(* IEC 61131-3 sources: traffic-lights/PLC_TrafficLights/Class/_OpenSSL (part 2) *)

	FUNCTION __CDECL VIRTUAL GLOBAL CRYPTO_add_lock
		VAR_INPUT
			pointer 	: ^DINT;
			amount 	: DINT;
			t 	: DINT;
			file 	: ^void;
			line 	: DINT;
		END_VAR
		VAR_OUTPUT
			RetVal (EAX) 	: DINT;
		END_VAR;

	FUNCTION GLOBAL TAB RetVal;
				//! <Function Comment="X509_LOOKUP_file is a certificate lookup method to use with X509_STORE, provided by OpenSSL library.&#13;&#10;&#13;&#10;The X509_LOOKUP_file method loads all the certificates or CRLs present in a file into memory at the time the file is added as a lookup source.&#13;&#10;&#13;&#10;File format is ASCII text which contains concatenated PEM certificates and CRLs.&#13;&#10;&#13;&#10;This method should be used by applications which work with a small set of CAs.&#13;&#10;&#13;&#10;See also www.openssl.org/docs/man1.1.0/crypto/X509_LOOKUP_file.html&#13;&#10;and       www.umich.edu/~x509/ssleay/x509_lookup.html&#13;&#10;and       www.umich.edu/~x509/ssleay/x509_store.html" Name="X509_LOOKUP_file"/>
	FUNCTION __CDECL VIRTUAL GLOBAL X509_LOOKUP_file
		VAR_OUTPUT
			RetAddr (EAX) 	: ^void;			//! <Variable Comment="X509_LOOKUP_file() returns a X509_LOOKUP_METHOD pointer to the static method x509_file_lookup(). &#13;&#10;This function is useful to call when you want to add a method to a stack of methods you are using. &#13;&#10;See X509_STORE documentation for more on this." Name="X509_LOOKUP_file.RetAddr"/>
		END_VAR;
				//! <Function Comment="Issues arbitrary control commands.&#13;&#10;&#13;&#10;See also www.openssl.org/docs/manmaster/man3/X509_LOOKUP_meth_set_get_by_fingerprint.html" Name="X509_LOOKUP_ctrl"/>
	FUNCTION __CDECL VIRTUAL GLOBAL X509_LOOKUP_ctrl
		VAR_INPUT
			ctx 	: ^void;			//! <Variable Comment="Pointer to X509_LOOKUP structure." Name="X509_LOOKUP_ctrl.ctx"/>
			cmd 	: DINT;			//! <Variable Comment="An arbitrary integer that defines some operation." Name="X509_LOOKUP_ctrl.cmd"/>
			argc 	: ^void;			//! <Variable Comment="Pointer to an array of characters.&#13;&#10;How argc and argl are used depends entirely on the control function." Name="X509_LOOKUP_ctrl.argc"/>
			argl 	: DINT;			//! <Variable Comment="Arbitrary integer.&#13;&#10;How argc and argl are used depends entirely on the control function." Name="X509_LOOKUP_ctrl.argl"/>
			retv 	: ^pVoid;			//! <Variable Comment="NULL or pointer to pointer to a location where any return data should be written to." Name="X509_LOOKUP_ctrl.retv"/>
		END_VAR
		VAR_OUTPUT
			RetVal (EAX) 	: DINT;			//! <Variable Comment="Returns -1 if no method table was found.&#13;&#10;              1 if no lookup method was found.&#13;&#10;" Name="X509_LOOKUP_ctrl.RetVal"/>
		END_VAR;
				//! <Function Comment="The X509_verify_cert() function attempts to discover and validate a certificate chain based on parameters in &lt;ctx&gt;. &#13;&#10;A complete description of the process is contained in the verify manual page. &#13;&#10;&#13;&#10;See also www.openssl.org/docs/manmaster/man3/X509_verify_cert.html" Name="X509_verify_cert"/>
	FUNCTION __CDECL VIRTUAL GLOBAL X509_verify_cert
		VAR_INPUT
			ctx 	: ^void;			//! <Variable Comment="Pointer to a context (X509_STORE_CTX structure)." Name="X509_verify_cert.ctx"/>
		END_VAR
		VAR_OUTPUT
			RetVal (EAX) 	: DINT;			//! <Variable Comment="If a complete chain can be built and validated this function returns 1, otherwise it return zero, in exceptional circumstances it can also return a negative code." Name="X509_verify_cert.RetVal"/>
		END_VAR;
				//! <Function Comment="X509_NAME_oneline() prints an ASCII version of &lt;a&gt; to &lt;buf&gt;. If &lt;buf&gt; is NULL then a buffer is dynamically allocated and returned, and &lt;size&gt; is ignored. &#13;&#10;Otherwise, at most &lt;size&gt; bytes will be written, including the ending &apos;\0&apos;, and &lt;buf&gt; is returned.&#13;&#10;&#13;&#10;NOTES&#13;&#10;X509_NAME_oneline() is a legacy function which produces a nonstandard output form, it doesn&apos;t handle multi character fields and has various quirks and inconsistencies. &#13;&#10;Its use is strongly discouraged in new applications.&#13;&#10;&#13;&#10;See also www.openssl.org/docs/man1.0.2/crypto/X509_NAME_oneline.html" Name="X509_NAME_oneline"/>
	FUNCTION __CDECL VIRTUAL GLOBAL X509_NAME_oneline
		VAR_INPUT
			a 	: ^void;			//! <Variable Comment="Pointer to a X509_NAME structure." Name="X509_NAME_oneline.a"/>
			buf 	: ^void;			//! <Variable Comment="Pointer to an output buffer or NULL (*char)." Name="X509_NAME_oneline.buf"/>
			size 	: DINT;			//! <Variable Comment="Output buffer size." Name="X509_NAME_oneline.size"/>
		END_VAR
		VAR_OUTPUT
			RetAddr (EAX) 	: ^void;			//! <Variable Comment="Pointer to the output buffer (*char)." Name="X509_NAME_oneline.RetAddr"/>
		END_VAR;
				//! <Function Comment="Internally loading of CRLs is implemented via function X509_load_crl_file. &#13;&#10;The function supports parameter &lt;typ&gt;, which can be one of constants FILETYPE_PEM, FILETYPE_ASN1 and FILETYPE_DEFAULT. &#13;&#10;It loads CRLs from specified &lt;file&gt; into memory cache of X509_STORE objects which given &lt;ctx&gt; parameter is associated with.&#13;&#10;&#13;&#10;See also www.openssl.org/docs/man1.1.0/crypto/X509_load_crl_file.html" Name="X509_load_crl_file"/>
	FUNCTION __CDECL VIRTUAL GLOBAL X509_load_crl_file
		VAR_INPUT
			ctx 	: ^void;			//! <Variable Comment="Pointer to X509_LOOKUP structure." Name="X509_load_crl_file.ctx"/>
			file 	: ^void;			//! <Variable Comment="Specifies the file to read from." Name="X509_load_crl_file.file"/>
			typ 	: DINT;			//! <Variable Comment="Can be one of constants FILETYPE_PEM, FILETYPE_ASN1 and FILETYPE_DEFAULT." Name="X509_load_crl_file.typ"/>
		END_VAR
		VAR_OUTPUT
			RetVal (EAX) 	: DINT;			//! <Variable Comment="Returns number of objects loaded from &lt;file&gt; or 0 in case of error." Name="X509_load_crl_file.RetVal"/>
		END_VAR;
				//! <Function Comment="X509_STORE_CTX_new() returns a newly initialised X509_STORE_CTX structure.&#13;&#10;&#13;&#10;NOTES&#13;&#10;The certificates and CRLs in a store are used internally and should not be freed up until after the associated X509_STORE_CTX is freed.&#13;&#10;&#13;&#10;BUGS&#13;&#10;The certificates and CRLs in a context are used internally and should not be freed up until after the associated X509_STORE_CTX is freed. &#13;&#10;Copies should be made, or reference counts increased instead.&#13;&#10;&#13;&#10;See also www.openssl.org/docs/man1.1.0/crypto/X509_STORE_CTX_new.html" Name="X509_STORE_CTX_new"/>
	FUNCTION __CDECL VIRTUAL GLOBAL X509_STORE_CTX_new
		VAR_OUTPUT
			RetAddr (EAX) 	: ^void;			//! <Variable Comment="Returns an newly allocated context (Pointer to X509_STORE_CTX structure) or &#13;&#10;NULL if an error occurred." Name="X509_STORE_CTX_new.RetAddr"/>
		END_VAR;
				//! <Function Comment="X509_STORE_CTX_free() completely frees up &lt;ctx&gt;. After this call &lt;ctx&gt; is no longer valid. &#13;&#10;If &lt;ctx&gt; is NULL nothing is done.&#13;&#10;&#13;&#10;See also www.openssl.org/docs/man1.1.0/crypto/X509_STORE_CTX_new.html" Name="X509_STORE_CTX_free"/>
	FUNCTION __CDECL VIRTUAL GLOBAL X509_STORE_CTX_free
		VAR_INPUT
			ctx 	: ^void;			//! <Variable Comment="Pointer to X509_STORE_CTX structure holding a context." Name="X509_STORE_CTX_free.ctx"/>
		END_VAR;
				//! <Function Comment="X509_STORE_CTX_init() sets up &lt;ctx&gt; for a subsequent verification operation. &#13;&#10;It must be called before each call to X509_verify_cert(), i.e. a &lt;ctx&gt; is only good for one call to X509_verify_cert(). &#13;&#10;If you want to verify a second certificate with the same &lt;ctx&gt; then you must call X509_STORE_CTX_cleanup() and then X509_STORE_CTX_init() again before the second call to X509_verify_cert(). &#13;&#10;The trusted certificate store is set to &lt;store&gt;, the end entity certificate to be verified is set to &lt;x509&gt; and a set of additional certificates (which will be untrusted but may be used to build the chain) in &lt;chain&gt;. &#13;&#10;Any or all of the &lt;store&gt;, &lt;x509&gt; and &lt;chain&gt; parameters can be NULL.&#13;&#10;&#13;&#10;See also www.openssl.org/docs/man1.1.0/crypto/X509_STORE_CTX_new.html" Name="X509_STORE_CTX_init"/>
	FUNCTION __CDECL VIRTUAL GLOBAL X509_STORE_CTX_init
		VAR_INPUT
			ctx 	: ^void;			//! <Variable Comment="Pointer to X509_STORE_CTX structure." Name="X509_STORE_CTX_init.ctx"/>
			store 	: ^void;			//! <Variable Comment="Pointer to X509_STORE structure or NULL" Name="X509_STORE_CTX_init.store"/>
			x509 	: ^void;			//! <Variable Comment="Pointer to X509 structure or NULL." Name="X509_STORE_CTX_init.x509"/>
			chain 	: ^void;			//! <Variable Comment="Pointer to STACK_OF(X509) or NULL." Name="X509_STORE_CTX_init.chain"/>
		END_VAR
		VAR_OUTPUT
			RetVal (EAX) 	: DINT;			//! <Variable Comment="Returns 1 for success or 0 if an error occurred." Name="X509_STORE_CTX_init.RetVal"/>
		END_VAR;
				//! <Function Comment="Returns the issuer name of certificate &lt;a&gt;. The returned value is an internal pointer which MUST NOT be freed.&#13;&#10;&#13;&#10;See also www.openssl.org/docs/man1.1.0/crypto/X509_get_subject_name.html" Name="X509_get_issuer_name"/>
	FUNCTION __CDECL VIRTUAL GLOBAL X509_get_issuer_name
		VAR_INPUT
			a 	: ^void;			//! <Variable Comment="Pointer to X509 structure holding a certificate." Name="X509_get_issuer_name.a"/>
		END_VAR
		VAR_OUTPUT
			RetAddr (EAX) 	: ^void;			//! <Variable Comment="Returns an X509_NAME pointer." Name="X509_get_issuer_name.RetAddr"/>
		END_VAR;
				//! <Function Comment="X509_LOOKUP_hash_dir is a certificate lookup method to use with X509_STORE, provided by OpenSSL library. &#13;&#10;X509_LOOKUP_hash_dir is a more advanced method, which loads certificates and CRLs on demand, and caches them in memory once they are loaded.&#13;&#10;&#13;&#10;See also www.openssl.org/docs/man1.1.0/crypto/X509_LOOKUP_hash_dir.html&#13;&#10;and       http://www.umich.edu/~x509/ssleay/x509_store.html" Name="X509_LOOKUP_hash_dir"/>
	FUNCTION __CDECL VIRTUAL GLOBAL X509_LOOKUP_hash_dir
		VAR_OUTPUT
			RetVal (EAX) 	: ^void;			//! <Variable Comment="Returns 1 on success or 0 on error. " Name="X509_LOOKUP_hash_dir.RetVal"/>
		END_VAR;
				//! <Function Comment="Sets the default values for the corresponding values used in certificate chain validation. &#13;&#10;Their behavior is documented in the corresponding X509_VERIFY_PARAM manual pages, e.g., X509_VERIFY_PARAM_set_depth(3).&#13;&#10;&#13;&#10;See also www.openssl.org/docs/manmaster/man3/X509_STORE_set_flags.html" Name="X509_STORE_set_flags"/>
	FUNCTION __CDECL VIRTUAL GLOBAL X509_STORE_set_flags
		VAR_INPUT
			ctx 	: ^void;			//! <Variable Comment="Pointer to X509_STORE structure.&#13;&#10;&#13;&#10;The X509_STORE structure is intended to be a consolidated mechanism for holding information about X.509 certificates and CRLs, and constructing and validating chains of certificates terminating in trusted roots. &#13;&#10;It admits multiple lookup mechanisms and efficient scaling performance with large numbers of certificates, and a great deal of flexibility in how validation and policy checks are performed." Name="X509_STORE_set_flags.ctx"/>
			flags 	: UDINT;			//! <Variable Comment="Flag values to set." Name="X509_STORE_set_flags.flags"/>
		END_VAR
		VAR_OUTPUT
			RetVal (EAX) 	: DINT;			//! <Variable Comment="Always returns 1, indicating success." Name="X509_STORE_set_flags.RetVal"/>
		END_VAR;
				//! <Function Comment="Adds the X509_LOOKUP_METHOD &lt;a&gt; to the stack &lt;v&gt;-&gt;get_cert_methods after creating an X509_LOOKUP that contains it as a subfield. &#13;&#10;It returns a pointer to the new X509_LOOKUP structure or NULL on error.&#13;&#10;&#13;&#10;X509_STORE_new() creates an empty X509_STORE structure, which contains no information about trusted certificates or where such certificates are located on disk, and is generally not usable. &#13;&#10;Normally, trusted certificates will be added to the X509_STORE to prepare it for use, via mechanisms such as X509_STORE_add_lookup() and X509_LOOKUP_file(), or PEM_read_bio_X509_AUX() &#13;&#10;and X509_STORE_add_cert(). &#13;&#10;CRLs can also be added, and many behaviors configured as desired.&#13;&#10;&#13;&#10;See also http://www.umich.edu/~x509/ssleay/x509_store.html&#13;&#10;" Name="X509_STORE_add_lookup"/>
	FUNCTION __CDECL VIRTUAL GLOBAL X509_STORE_add_lookup
		VAR_INPUT
			v 	: ^void;			//! <Variable Comment="Pointer to X509_STORE structure." Name="X509_STORE_add_lookup.v"/>
			a 	: ^void;			//! <Variable Comment="Pointer to X509_LOOKUP_METHOD structure holding a lookup method." Name="X509_STORE_add_lookup.a"/>
		END_VAR
		VAR_OUTPUT
			RetAddr (EAX) 	: ^void;			//! <Variable Comment="Returns a pointer to the new X509_LOOKUP structure or NULL on error." Name="X509_STORE_add_lookup.RetAddr"/>
		END_VAR;
				//! <Function Comment="X509_STORE_set_default_paths() is somewhat misnamed, in that it does not set what default paths should be used for loading certificates. &#13;&#10;Instead, it loads certificates into the X509_STORE from the hardcoded default paths.&#13;&#10;&#13;&#10;See also www.openssl.org/docs/man1.1.1/man3/X509_STORE_set_default_paths.html&#13;&#10;and       http://www.umich.edu/~x509/ssleay/x509_store.html" Name="X509_STORE_set_default_paths"/>
	FUNCTION __CDECL VIRTUAL GLOBAL X509_STORE_set_default_paths
		VAR_INPUT
			ctx 	: ^void;			//! <Variable Comment="Pointer to X509_STORE structure." Name="X509_STORE_set_default_paths.ctx"/>
		END_VAR
		VAR_OUTPUT
			RetVal (EAX) 	: DINT;			//! <Variable Comment="Returns 1 on success or 0 on failure." Name="X509_STORE_set_default_paths.RetVal"/>
		END_VAR;
				//! <Function Comment="Is used to retrieve application specific data. Returns the application data or 0 on failure. &#13;&#10;0 may also be valid application data but currently it can only fail if given an invalid &lt;idx&gt; parameter.&#13;&#10;&#13;&#10;See also www.openssl.org/docs/man1.0.2/crypto/X509_STORE_CTX_get_ex_data.html&#13;&#10;and       www.openssl.org/docs/man1.0.2/crypto/RSA_get_ex_new_index.html" Name="X509_STORE_CTX_get_ex_data"/>
	FUNCTION __CDECL VIRTUAL GLOBAL X509_STORE_CTX_get_ex_data
		VAR_INPUT
			ctx 	: ^void;			//! <Variable Comment="Pointer to X509_STORE_CTX structure." Name="X509_STORE_CTX_get_ex_data.ctx"/>
			idx 	: DINT;			//! <Variable Comment="Index retrieved by RSA_get_ex_new_index()." Name="X509_STORE_CTX_get_ex_data.idx"/>
		END_VAR
		VAR_OUTPUT
			RetAddr (EAX) 	: ^void;			//! <Variable Comment="Pointer to the retrieved application data or NULL on failure.&#13;&#10;Since the application data can be anything at all it is passed and retrieved as a void * type." Name="X509_STORE_CTX_get_ex_data.RetAddr"/>
		END_VAR;
				//! <Function Comment="Is used to set application specific data, the data is supplied in the &lt;data&gt; parameter and its precise meaning is up to the application.&#13;&#10;&#13;&#10;See also www.openssl.org/docs/man1.0.2/crypto/X509_STORE_CTX_get_ex_data.html&#13;&#10;and       www.openssl.org/docs/man1.0.2/crypto/RSA_get_ex_new_index.html" Name="X509_STORE_CTX_set_ex_data"/>
	FUNCTION __CDECL VIRTUAL GLOBAL X509_STORE_CTX_set_ex_data
		VAR_INPUT
			ctx 	: ^void;			//! <Variable Comment="Pointer to X509_STORE_CTX structure." Name="X509_STORE_CTX_set_ex_data.ctx"/>
			idx 	: DINT;			//! <Variable Comment="Index retrieved by RSA_get_ex_new_index()." Name="X509_STORE_CTX_set_ex_data.idx"/>
			data 	: ^void;			//! <Variable Comment="Pointer to the application data.&#13;&#10;Since the application data can be anything at all it is passed as a void * type." Name="X509_STORE_CTX_set_ex_data.data"/>
		END_VAR
		VAR_OUTPUT
			RetVal (EAX) 	: DINT;			//! <Variable Comment="Returns 1 on success or 0 on failure." Name="X509_STORE_CTX_set_ex_data.RetVal"/>
		END_VAR;
				//! <Function Comment="X509_STORE_CTX_get_error() returns the error code of &lt;ctx&gt;, see the ERROR CODES section for a full description of all error codes. &#13;&#10;&#13;&#10;This function is typically called after X509_verify_cert() has indicated an error or in a verification callback to determine the nature of an error.&#13;&#10;&#13;&#10;See also www.openssl.org/docs/man1.0.2/crypto/X509_STORE_CTX_get_error.html" Name="X509_STORE_CTX_get_error"/>
	FUNCTION __CDECL VIRTUAL GLOBAL X509_STORE_CTX_get_error
		VAR_INPUT
			ctx 	: ^void;			//! <Variable Comment="Pointer to X509_STORE_CTX structure." Name="X509_STORE_CTX_get_error.ctx"/>
		END_VAR
		VAR_OUTPUT
			RetVal (EAX) 	: DINT;			//! <Variable Comment="Returns X509_V_OK or an error code.&#13;&#10;&#13;&#10;See the class documentation for a list of error codes and messages." Name="X509_STORE_CTX_get_error.RetVal"/>
		END_VAR;
				//! <Function Comment="X509_STORE_CTX_get_current_cert() returns the certificate in &lt;ctx&gt; which caused the error or NULL if no certificate is relevant.&#13;&#10;&#13;&#10;This function is typically called after X509_verify_cert() has indicated an error or in a verification callback to determine the nature of an error.&#13;&#10;&#13;&#10;See also www.openssl.org/docs/man1.0.2/crypto/X509_STORE_CTX_get_error.html" Name="X509_STORE_CTX_get_current_cert"/>
	FUNCTION __CDECL VIRTUAL GLOBAL X509_STORE_CTX_get_current_cert
		VAR_INPUT
			ctx 	: ^void;			//! <Variable Comment="Pointer to X509_STORE_CTX structure." Name="X509_STORE_CTX_get_current_cert.ctx"/>
		END_VAR
		VAR_OUTPUT
			RetAddr (EAX) 	: ^void;			//! <Variable Comment="Returns a X509 pointer to the certificate which caused the error or NULL if no certificate is relevant to the error." Name="X509_STORE_CTX_get_current_cert.RetAddr"/>
		END_VAR;
				//! <Function Comment="X509_STORE_CTX_get_error_depth() returns the depth of the error. This is a non-negative integer representing where in the certificate chain the error occurred. &#13;&#10;If it is zero it occurred in the end entity certificate, one if it is the certificate which signed the end entity certificate and so on.&#13;&#10;&#13;&#10;This function is typically called after X509_verify_cert() has indicated an error or in a verification callback to determine the nature of an error.&#13;&#10;&#13;&#10;See also www.openssl.org/docs/man1.0.2/crypto/X509_STORE_CTX_get_error.html" Name="X509_STORE_CTX_get_error_depth"/>
	FUNCTION __CDECL VIRTUAL GLOBAL X509_STORE_CTX_get_error_depth
		VAR_INPUT
			ctx 	: ^void;			//! <Variable Comment="Pointer to X509_STORE_CTX structure." Name="X509_STORE_CTX_get_error_depth.ctx"/>
		END_VAR
		VAR_OUTPUT
			RetVal (EAX) 	: DINT;			//! <Variable Comment="Returns a non-negative error depth." Name="X509_STORE_CTX_get_error_depth.RetVal"/>
		END_VAR;
				//! <Function Comment="X509_verify_cert_error_string() returns a human readable error string for verification of error &lt;a&gt;." Name="X509_verify_cert_error_string"/>
	FUNCTION __CDECL VIRTUAL GLOBAL X509_verify_cert_error_string
		VAR_INPUT
			a 	: DINT;			//! <Variable Comment="Error number." Name="X509_verify_cert_error_string.a"/>
		END_VAR
		VAR_OUTPUT
			RetAddr (EAX) 	: ^void;			//! <Variable Comment="Returns a human readable error string for verification of error &lt;a&gt;." Name="X509_verify_cert_error_string.RetAddr"/>
		END_VAR;
				//! <Function Comment="i2d_PublicKey() encodes key &lt;a&gt; into DER format. It uses a key specific format or, if none is defined for that key type, PKCS#8 unencrypted PublicKeyInfo format.&#13;&#10;&#13;&#10;NOTES&#13;&#10;The EVP_PKEY structure passed to the function should have all the public key components present.&#13;&#10;&#13;&#10;The encoded data is in binary form and may contain embedded zeroes. Functions such as strlen() will not return the correct length of the encoded structure.&#13;&#10;&#13;&#10;See also www.openssl.org/docs/man1.1.0/crypto/i2d_PublicKey.html&#13;&#10;and       www.openssl.org/docs/man1.0.2/crypto/i2d_RSAPublicKey.html&#13;&#10;and       www.openssl.org/docs/manmaster/man3/i2d_RSA_PUBKEY.html" Name="i2d_PublicKey"/>
	FUNCTION __CDECL VIRTUAL GLOBAL i2d_PublicKey
		VAR_INPUT
			a 	: ^void;			//! <Variable Comment="Pointer to a EVP_PKEY structure holding the public key." Name="i2d_PublicKey.a"/>
			pp 	: ^pVoid;			//! <Variable Comment="Pointer to pointer to output buffer (i.e. **char).&#13;&#10;If &lt;pp&gt; is not NULL, the DER encoded data is written to the buffer at *&lt;pp&gt;, and *&lt;pp&gt; is incremented to point after the data just written.&#13;&#10;If *&lt;pp&gt; is NULL memory will be allocated for a buffer and the encoded data written to it. In this case *&lt;pp&gt; is not incremented and it points to the start of the data just written." Name="i2d_PublicKey.pp"/>
		END_VAR
		VAR_OUTPUT
			RetVal (EAX) 	: DINT;			//! <Variable Comment="Returns the number of bytes successfully encoded or a negative value if an error occurs. &#13;&#10;The error code can be obtained by calling ERR_get_error()." Name="i2d_PublicKey.RetVal"/>
		END_VAR;
				//! <Function Comment="EVP_PKEY_type() returns the type of key corresponding to the value &lt;typ&gt;. &#13;&#10;The type of a key can be obtained with EVP_PKEY_type(pkey-&gt;type). &#13;&#10;&#13;&#10;See also www.openssl.org/docs/man1.0.2/crypto/EVP_PKEY_type.html" Name="EVP_PKEY_type"/>
	FUNCTION __CDECL VIRTUAL GLOBAL EVP_PKEY_type
		VAR_INPUT
			typ 	: DINT;			//! <Variable Comment="Value retrieved with pkey-&gt;type." Name="EVP_PKEY_type.typ"/>
		END_VAR
		VAR_OUTPUT
			RetVal (EAX) 	: DINT;			//! <Variable Comment="The return value will be EVP_PKEY_RSA, EVP_PKEY_DSA, EVP_PKEY_DH or EVP_PKEY_EC for the corresponding key types or NID_undef if the key type is unassigned." Name="EVP_PKEY_type.RetVal"/>
		END_VAR;
				//! <Function Comment="Do not use this function in new code. It is provided purely for compatibility with legacy application code.&#13;&#10;This function is a wrapper around the corresponding standard realloc() function.&#13;&#10;&#13;&#10;See also www.openssl.org/docs/man1.1.0/crypto/CRYPTO_realloc.html&#13;&#10;and       http://man.openbsd.org/OpenBSD-6.1/OPENSSL_realloc.3" Name="CRYPTO_realloc"/>
	FUNCTION __CDECL VIRTUAL GLOBAL CRYPTO_realloc
		VAR_INPUT
			addr 	: ^void;			//! <Variable Comment="Pointer to a memory block previously allocated." Name="CRYPTO_realloc.addr"/>
			num 	: DINT;			//! <Variable Comment="New size for the memory block, in bytes." Name="CRYPTO_realloc.num"/>
			file 	: ^void;			//! <Variable Comment="The Structured Text __FILE__ parameter." Name="CRYPTO_realloc.file"/>
			line 	: DINT;			//! <Variable Comment="The Structured Text __LINE__ parameter." Name="CRYPTO_realloc.line"/>
		END_VAR
		VAR_OUTPUT
			RetAddr (EAX) 	: ^void;			//! <Variable Comment="Returns a void pointer to allocated memory or NULL on error." Name="CRYPTO_realloc.RetAddr"/>
		END_VAR;
				//! <Function Comment="BIO_ctrl() is a BIO &quot;control&quot; operation taking arguments of various types. &#13;&#10;This function is not normally called directly, various macros are used instead. &#13;&#10;The standard macros are described below, macros specific to a particular type of BIO are described in the specific BIOs manual page as well as any special features of the standard calls.&#13;&#10;&#13;&#10;A BIO is an I/O abstraction, it hides many of the underlying I/O details from an application. &#13;&#10;If an application uses a BIO for its I/O it can transparently handle SSL connections, unencrypted network connections and file I/O.&#13;&#10;&#13;&#10;See also www.openssl.org/docs/man1.0.2/crypto/BIO_ctrl.html&#13;&#10;and       www.openssl.org/docs/man1.0.2/crypto/BIO_get_read_request.html&#13;&#10;and       www.openssl.org/docs/man1.0.2/crypto/BIO_new_buffer_ssl_connect.html&#13;&#10;and       www.openssl.org/docs/man1.0.2/crypto/BIO_ctrl_reset_read_request.html&#13;&#10;and       www.openssl.org/docs/man1.0.2/crypto/BIO_f_buffer.html&#13;&#10;and       www.openssl.org/docs/man1.0.2/crypto/BIO_set_fd.html&#13;&#10;and       www.openssl.org/docs/man1.1.1/man7/bio.html" Name="BIO_ctrl"/>
	FUNCTION __CDECL VIRTUAL GLOBAL BIO_ctrl
		VAR_INPUT
			b 	: ^void;			//! <Variable Comment="Pointer to BIO structure." Name="BIO_ctrl.b"/>
			cmd 	: DINT;			//! <Variable Comment="Command code.&#13;&#10;E.g. BIO_C_MAKE_BIO_PAIR, BIO_C_DESTROY_BIO_PAIR, &#13;&#10;BIO_C_SHUTDOWN_WR, BIO_C_SET_WRITE_BUF_SIZE, BIO_C_GET_WRITE_BUF_SIZE, &#13;&#10;BIO_C_GET_WRITE_GUARANTEE, BIO_C_GET_READ_REQUEST,&#13;&#10;BIO_C_SET_SSL, BIO_C_GET_SSL,&#13;&#10;BIO_C_SSL_MODE,&#13;&#10;BIO_C_SET_SSL_RENEGOTIATE_BYTES,&#13;&#10;BIO_C_SET_SSL_RENEGOTIATE_TIMEOUT,&#13;&#10;BIO_C_SET_SSL_NUM_RENEGOTIATES,&#13;&#10;BIO_C_DO_STATE_MACHINE ........" Name="BIO_ctrl.cmd"/>
			larg 	: DINT;			//! <Variable Comment="The meaning of &lt;larg&gt; depends on parameter &lt;cmd&gt;." Name="BIO_ctrl.larg"/>
			parg 	: ^void;			//! <Variable Comment="The meaning of &lt;parg&gt; depends on parameter &lt;cmd&gt;." Name="BIO_ctrl.parg"/>
		END_VAR
		VAR_OUTPUT
			RetVal (EAX) 	: DINT;			//! <Variable Comment="The meaning of &lt;RetVal&gt; depends on parameter &lt;cmd&gt;." Name="BIO_ctrl.RetVal"/>
		END_VAR;
				//! <Function Comment="BIO_s_mem() returns the memory BIO method function.&#13;&#10;A memory BIO is a source/sink BIO which uses memory for its I/O." Name="BIO_s_mem"/>
	FUNCTION __CDECL VIRTUAL GLOBAL BIO_s_mem
		VAR_OUTPUT
			RetAddr (EAX) 	: ^void;			//! <Variable Comment="Returns a BIO_METHOD pointer to the memory BIO method function." Name="BIO_s_mem.RetAddr"/>
		END_VAR;
				//! <Function Comment="BIO_s_file() returns the BIO file method. As its name implies it is a wrapper round the stdio FILE structure and it is a source/sink BIO.&#13;&#10;&#13;&#10;See also www.openssl.org/docs/man1.0.2/crypto/BIO_s_file.html" Name="BIO_s_file"/>
	FUNCTION __CDECL VIRTUAL GLOBAL BIO_s_file
		VAR_OUTPUT
			RetAddr (EAX) 	: ^void;			//! <Variable Comment="Returns a BIO_METHOD pointer to the BIO file method." Name="BIO_s_file.RetAddr"/>
		END_VAR;
				//! <Function Comment="X509_get_ext() operates on the extensions of certificate &lt;x&gt;. It is otherwise identical to X509v3_get_ext().&#13;&#10;&#13;&#10;X509v3_get_ext() retrieves extension &lt;loc&gt; from &lt;x&gt;. The index &lt;loc&gt; can take any value from 0 to X509_get_ext_count(&lt;x&gt;) - 1. &#13;&#10;The returned extension is an internal pointer which must not be freed up by the application.&#13;&#10;&#13;&#10;See also www.openssl.org/docs/man1.1.0/crypto/X509_get_ext.html" Name="X509_get_ext"/>
	FUNCTION __CDECL VIRTUAL GLOBAL X509_get_ext
		VAR_INPUT
			x 	: ^void;			//! <Variable Comment="Pointer to X509 structure holding a certificate." Name="X509_get_ext.x"/>
			loc 	: DINT;			//! <Variable Comment="Any value from 0 to X509_get_ext_count(&lt;x&gt;) - 1. " Name="X509_get_ext.loc"/>
		END_VAR
		VAR_OUTPUT
			RetAddr (EAX) 	: ^void;			//! <Variable Comment="Returns an X509_EXTENSION pointer or NULL if an error occurs." Name="X509_get_ext.RetAddr"/>
		END_VAR;
				//! <Function Comment="The function EVP_PKEY_cmp() compares the public key components and parameters (if present) of keys &lt;a&gt; and &lt;b&gt;.&#13;&#10;&#13;&#10;See also www.openssl.org/docs/man1.0.2/crypto/EVP_PKEY_cmp.html" Name="EVP_PKEY_cmp"/>
	FUNCTION __CDECL VIRTUAL GLOBAL EVP_PKEY_cmp
		VAR_INPUT
			a 	: ^void;			//! <Variable Comment="EVP_PKEY pointer to first key." Name="EVP_PKEY_cmp.a"/>
			b 	: ^void;			//! <Variable Comment="EVP_PKEY pointer to second key." Name="EVP_PKEY_cmp.b"/>
		END_VAR
		VAR_OUTPUT
			RetVal (EAX) 	: DINT;			//! <Variable Comment="Returns &#13;&#10;1 if the keys match, &#13;&#10;0 if they don&apos;t match, &#13;&#10;-1 if the key types are different and &#13;&#10;-2 if the operation is not supported." Name="EVP_PKEY_cmp.RetVal"/>
		END_VAR;
				//! <Function Comment="The EVP_PKEY_new() function allocates an empty EVP_PKEY structure which is used by OpenSSL to store private keys.&#13;&#10;EVP_PKEY_free() frees up the private key key.&#13;&#10;&#13;&#10;NOTES&#13;&#10;The EVP_PKEY structure is used by various OpenSSL functions which require a general private key without reference to any particular algorithm.&#13;&#10;&#13;&#10;The structure returned by EVP_PKEY_new() is empty. To add a private key to this empty structure the functions described in EVP_PKEY_set1_RSA should be used.&#13;&#10;&#13;&#10;See also www.openssl.org/docs/man1.0.2/crypto/EVP_PKEY_new.html" Name="EVP_PKEY_new"/>
	FUNCTION __CDECL VIRTUAL GLOBAL EVP_PKEY_new
		VAR_OUTPUT
			RetAddr (EAX) 	: ^void;			//! <Variable Comment="Returns either a pointer to the newly allocated EVP_PKEY structure of NULL if an error occurred." Name="EVP_PKEY_new.RetAddr"/>
		END_VAR;
				//! <Function Comment="The function ASN1_TIME_set() sets the ASN1_TIME structure &lt;sx&gt; to the time represented by the time_t value &lt;tx&gt;. &#13;&#10;If &lt;sx&gt; is NULL a new ASN1_TIME structure is allocated and returned.&#13;&#10;&#13;&#10;See also www.openssl.org/docs/man1.0.2/crypto/ASN1_TIME_set.html" Name="ASN1_TIME_set"/>
	FUNCTION __CDECL VIRTUAL GLOBAL ASN1_TIME_set
		VAR_INPUT
			sx 	: ^void;			//! <Variable Comment="Pointer to ASN1_TIME structure.&#13;&#10;&lt;sx&gt; must satisfy the ASN1_TIME format mandated by RFC 5280, i.e., its format must be either YYMMDDHHMMSSZ or YYYYMMDDHHMMSSZ (it&apos;s a literal Z at the end, meaning &quot;Zulu&quot;).&#13;&#10;" Name="ASN1_TIME_set.sx"/>
			tx 	: DINT;			//! <Variable Comment="Number of seconds since the start of the Unix epoch: midnight UTC of January 1, 1970 (not counting leap seconds)." Name="ASN1_TIME_set.tx"/>
		END_VAR
		VAR_OUTPUT
			RetAddr (EAX) 	: ^void;			//! <Variable Comment="Returns a pointer to an ASN1_TIME structure or NULL if an error occurred." Name="ASN1_TIME_set.RetAddr"/>
		END_VAR;
				//! <Function Comment="X509_CRL_sign() signs CRLs (Certificate Revocation Lists).&#13;&#10;&#13;&#10;See also www.openssl.org/docs/man1.1.0/crypto/X509_CRL_sign.html" Name="X509_CRL_sign"/>
	FUNCTION __CDECL VIRTUAL GLOBAL X509_CRL_sign
		VAR_INPUT
			x 	: ^void;			//! <Variable Comment="Pointer to X509_CRL structure holding a certificate revocation list (CRL)." Name="X509_CRL_sign.x"/>
			pkey 	: ^void;			//! <Variable Comment="Pointer to a EVP_PKEY structure holding the private key." Name="X509_CRL_sign.pkey"/>
			md 	: ^void;			//! <Variable Comment="Pointer to a EVP_MD structure holding the message digest." Name="X509_CRL_sign.md"/>
		END_VAR
		VAR_OUTPUT
			RetVal (EAX) 	: DINT;			//! <Variable Comment="Returns the size of the signature in bytes for success and zero for failure." Name="X509_CRL_sign.RetVal"/>
		END_VAR;
				//! <Function Comment="X509_PUBKEY_get() returns the public key contained in &lt;key&gt;.&#13;&#10;The reference count on the returned key is incremented so it MUST be freed using EVP_PKEY_free() after use.&#13;&#10;&#13;&#10;See also www.openssl.org/docs/man1.1.0/crypto/i2d_PUBKEY.html" Name="X509_PUBKEY_get"/>
	FUNCTION __CDECL VIRTUAL GLOBAL X509_PUBKEY_get
		VAR_INPUT
			key 	: ^void;			//! <Variable Comment="Pointer to a X509_PUBKEY structure." Name="X509_PUBKEY_get.key"/>
		END_VAR
		VAR_OUTPUT
			RetAddr (EAX) 	: ^void;			//! <Variable Comment="Returns a pointer to an EVP_PKEY structure or NULL if an error occurs." Name="X509_PUBKEY_get.RetAddr"/>
		END_VAR;
				//! <Function Comment="Sets the referenced &lt;pkey&gt; to &lt;key&gt; however it uses the supplied &lt;key&gt; internally and so &lt;key&gt; will be freed when the parent &lt;pkey&gt; is freed.&#13;&#10;&#13;&#10;See also www.openssl.org/docs/manmaster/man3/EVP_PKEY_set1_RSA.html" Name="EVP_PKEY_assign"/>
	FUNCTION __CDECL VIRTUAL GLOBAL EVP_PKEY_assign
		VAR_INPUT
			pKey 	: ^void;			//! <Variable Comment="Pointer to a EVP_PKEY structure." Name="EVP_PKEY_assign.pKey"/>
			typ 	: DINT;			//! <Variable Comment="Type of &lt;pkey&gt;.&#13;&#10;EVP_PKEY_RSA, EVP_PKEY_DSA, EVP_PKEY_DH or EVP_PKEY_EC." Name="EVP_PKEY_assign.typ"/>
			key 	: ^void;			//! <Variable Comment="Void pointer to the key data." Name="EVP_PKEY_assign.key"/>
		END_VAR
		VAR_OUTPUT
			RetVal (EAX) 	: DINT;			//! <Variable Comment="Returns 1 for success and 0 for failure." Name="EVP_PKEY_assign.RetVal"/>
		END_VAR;
				//! <Function Comment="This function prints out an individual extension to a BIO pointer." Name="X509V3_EXT_print"/>
	FUNCTION __CDECL VIRTUAL GLOBAL X509V3_EXT_print
		VAR_INPUT
			out 	: ^void;			//! <Variable Comment="BIO pointer to which the extension is printed." Name="X509V3_EXT_print.out"/>
			ext 	: ^void;			//! <Variable Comment="Pointer to the X509_EXTENSION that will be printed to &lt;out&gt;." Name="X509V3_EXT_print.ext"/>
			flag 	: UDINT;			//! <Variable Comment="Currently the &lt;flag&gt; argument is unused and should be set to 0." Name="X509V3_EXT_print.flag"/>
			indent 	: DINT;			//! <Variable Comment="&lt;indent&gt; is the number of spaces to indent each line.&#13;&#10;" Name="X509V3_EXT_print.indent"/>
		END_VAR
		VAR_OUTPUT
			RetVal (EAX) 	: DINT;			//! <Variable Comment="Returns 1 for success and 0 for failure." Name="X509V3_EXT_print.RetVal"/>
		END_VAR;
				//! <Function Comment="X509_get_ext_by_NID() looks for an extension with &lt;nid&gt; from certificate &lt;x&gt;. &#13;&#10;The search starts from the extension after &lt;lastpos&gt; or from the beginning if &lt;lastpos&gt; is -1. If the extension is found its index is returned otherwise -1 is returned.&#13;&#10;&#13;&#10;See also www.openssl.org/docs/man1.1.0/crypto/X509_REVOKED_get_ext.html" Name="X509_get_ext_by_NID"/>
	FUNCTION __CDECL VIRTUAL GLOBAL X509_get_ext_by_NID
		VAR_INPUT
			x 	: ^void;			//! <Variable Comment="Pointer to a X509 structure holding a certificate." Name="X509_get_ext_by_NID.x"/>
			nid 	: DINT;			//! <Variable Comment="NID value." Name="X509_get_ext_by_NID.nid"/>
			lastpos 	: DINT;			//! <Variable Comment="Should initially be set to -1, if it is set to zero the initial extension will not be checked." Name="X509_get_ext_by_NID.lastpos"/>
		END_VAR
		VAR_OUTPUT
			RetVal (EAX) 	: DINT;			//! <Variable Comment="Returns the extension index or -1 if an error occurs.&#13;&#10;Extension indices start from zero, so a zero index return value is not an error." Name="X509_get_ext_by_NID.RetVal"/>
		END_VAR;
				//! <Function Comment="Sets the version number of a CRL (Certificate Revocation List).&#13;&#10;&#13;&#10;NOTES&#13;&#10;The version field of certificates, certificate requests and CRLs has a DEFAULT value of v1(0) meaning the field should be omitted for version 1. &#13;&#10;This is handled transparently by this function.&#13;&#10;&#13;&#10;See also www.openssl.org/docs/man1.1.0/crypto/X509_CRL_set_version.html" Name="X509_CRL_set_version"/>
	FUNCTION __CDECL VIRTUAL GLOBAL X509_CRL_set_version
		VAR_INPUT
			x 	: ^void;			//! <Variable Comment="Pointer to X509_CRL structure holding a certificate revocation list (CRL)." Name="X509_CRL_set_version.x"/>
			version 	: DINT;			//! <Variable Comment="Version number." Name="X509_CRL_set_version.version"/>
		END_VAR
		VAR_OUTPUT
			RetVal (EAX) 	: DINT;			//! <Variable Comment="Returns 1 for success and 0 for failure." Name="X509_CRL_set_version.RetVal"/>
		END_VAR;
				//! <Function Comment="X509_CRL_add0_revoked() appends revoked entry &lt;rev&gt; to CRL &lt;crl&gt;. &#13;&#10;The pointer &lt;rev&gt; is used internally so it must not be freed up after the call: it is freed when the parent CRL is freed.&#13;&#10;&#13;&#10;See also www.openssl.org/docs/man1.1.0/crypto/X509_CRL_add0_revoked.html&#13;&#10;and        www.openssl.org/docs/man1.0.2/crypto/crypto.html" Name="X509_CRL_add0_revoked"/>
	FUNCTION __CDECL VIRTUAL GLOBAL X509_CRL_add0_revoked
		VAR_INPUT
			crl 	: ^void;			//! <Variable Comment="Pointer to X509_CRL structure holding a certificate revocation list (CRL)." Name="X509_CRL_add0_revoked.crl"/>
			rev 	: ^void;			//! <Variable Comment="Pointer to a X509_REVOKED structure holding the revoked entry." Name="X509_CRL_add0_revoked.rev"/>
		END_VAR
		VAR_OUTPUT
			RetVal (EAX) 	: DINT;			//! <Variable Comment="Returns 1 for success and 0 for failure." Name="X509_CRL_add0_revoked.RetVal"/>
		END_VAR;
				//! <Function Comment="X509_CRL_add1_ext_i2d() adds extension &lt;value&gt; to CRL &lt;x&gt; using OID &lt;nid&gt; and criticality &lt;crit&gt; according to &lt;flags&gt;.&#13;&#10;&#13;&#10;See also www.openssl.org/docs/man1.1.0/crypto/X509_CRL_add1_ext_i2d.html" Name="X509_CRL_add1_ext_i2d"/>
	FUNCTION __CDECL VIRTUAL GLOBAL X509_CRL_add1_ext_i2d
		VAR_INPUT
			x 	: ^void;			//! <Variable Comment="Pointer to X509_CRL structure holding a certificate revocation list (CRL)." Name="X509_CRL_add1_ext_i2d.x"/>
			nid 	: DINT;			//! <Variable Comment="NID (Numeric Identifier) value." Name="X509_CRL_add1_ext_i2d.nid"/>
			value 	: ^void;			//! <Variable Comment="Void pointer to the extension data to be added." Name="X509_CRL_add1_ext_i2d.value"/>
			crit 	: DINT;			//! <Variable Comment="Determines the value of X509_EXTENSION.critical.&#13;&#10;0 if the extension is not critical.&#13;&#10;1 if the extension is critical." Name="X509_CRL_add1_ext_i2d.crit"/>
			flags 	: UDINT;			//! <Variable Comment="The &lt;flags&gt; parameter may be one of the following values.&#13;&#10;&#13;&#10;X509V3_ADD_DEFAULT appends a new extension only if the extension does not already exist. An error is returned if the extension does already exist.&#13;&#10;&#13;&#10;X509V3_ADD_APPEND appends a new extension, ignoring whether the extension already exists.&#13;&#10;&#13;&#10;X509V3_ADD_REPLACE replaces an extension if it exists otherwise appends a new extension.&#13;&#10;&#13;&#10;X509V3_ADD_REPLACE_EXISTING replaces an existing extension if it exists otherwise returns an error.&#13;&#10;&#13;&#10;X509V3_ADD_KEEP_EXISTING appends a new extension only if the extension does not already exist. An error is not returned if the extension does already exist.&#13;&#10;&#13;&#10;X509V3_ADD_DELETE extension nid is deleted: no new extension is added.&#13;&#10;&#13;&#10;If X509V3_ADD_SILENT is ored with flags: any error returned will not be added to the error queue." Name="X509_CRL_add1_ext_i2d.flags"/>
		END_VAR
		VAR_OUTPUT
			RetVal (EAX) 	: DINT;			//! <Variable Comment="Returns &#13;&#10;1 if the operation is successful and &#13;&#10;0 if it fails due to a non-fatal error (extension not found, already exists, cannot be encoded) or &#13;&#10;-1 due to a fatal error such as a memory allocation failure." Name="X509_CRL_add1_ext_i2d.RetVal"/>
		END_VAR;
				//! <Function Comment="Together with X509_CRL_set_nextUpdate() it sets the validity period of the CRL &lt;x&gt;.&#13;&#10;&#13;&#10;See also https://metacpan.org/pod/Crypt::OpenSSL::CA#set_lastUpdate-($enddate)" Name="X509_CRL_set_lastUpdate"/>
	FUNCTION __CDECL VIRTUAL GLOBAL X509_CRL_set_lastUpdate
		VAR_INPUT
			x 	: ^void;			//! <Variable Comment="Pointer to X509_CRL structure holding a certificate revocation list (CRL)." Name="X509_CRL_set_lastUpdate.x"/>
			tm 	: ^void;			//! <Variable Comment="Pointer to ASN1_TIME structure holding the enddate.&#13;&#10;The date must be in the GMT timezone, with the format yyyymmddhhmmssZ (it&apos;s a literal Z at the end, meaning &quot;Zulu&quot;)." Name="X509_CRL_set_lastUpdate.tm"/>
		END_VAR
		VAR_OUTPUT
			RetVal (EAX) 	: DINT;			//! <Variable Comment="Returns 1 for success of 0 if an error occurred." Name="X509_CRL_set_lastUpdate.RetVal"/>
		END_VAR;
				//! <Function Comment="Together with X509_CRL_set_lastUpdate() it sets the validity period of the CRL &lt;x&gt;.&#13;&#10;&#13;&#10;See also https://metacpan.org/pod/Crypt::OpenSSL::CA#set_lastUpdate-($enddate)" Name="X509_CRL_set_nextUpdate"/>
	FUNCTION __CDECL VIRTUAL GLOBAL X509_CRL_set_nextUpdate
		VAR_INPUT
			x 	: ^void;			//! <Variable Comment="Pointer to X509_CRL structure holding a certificate revocation list (CRL)." Name="X509_CRL_set_nextUpdate.x"/>
			tm 	: ^void;			//! <Variable Comment="Pointer to ASN1_TIME structure holding the startdate.&#13;&#10;The date must be in the GMT timezone, with the format yyyymmddhhmmssZ (it&apos;s a literal Z at the end, meaning &quot;Zulu&quot;)." Name="X509_CRL_set_nextUpdate.tm"/>
		END_VAR
		VAR_OUTPUT
			RetVal (EAX) 	: DINT;			//! <Variable Comment="Returns 1 for success of 0 if an error occurred." Name="X509_CRL_set_nextUpdate.RetVal"/>
		END_VAR;
				//! <Function Comment="Add a field whose name is defined by the string &lt;field&gt; to &lt;name&gt;. The field value to be added is in &lt;bytes&gt; of length &lt;len&gt;. &#13;&#10;If &lt;len&gt; is -1 then the field length is calculated internally using strlen(&lt;bytes&gt;).&#13;&#10;&#13;&#10;The type of field is determined by &lt;typ&gt; which can either be a definition of the type of bytes (such as MBSTRING_ASC) or a standard ASN1 type (such as V_ASN1_IA5STRING). &#13;&#10;&#13;&#10;The &lt;loc&gt; and &lt;set&gt; parameters determine where a new entry should be added. For almost all applications &lt;loc&gt; can be set to -1 and &lt;set&gt; to 0. &#13;&#10;This adds a new entry to the end of &lt;name&gt; as a single valued RelativeDistinguishedName (RDN).&#13;&#10;&#13;&#10;See also www.openssl.org/docs/man1.1.0/crypto/X509_NAME_add_entry_by_txt.html" Name="X509_NAME_add_entry_by_txt"/>
	FUNCTION __CDECL VIRTUAL GLOBAL X509_NAME_add_entry_by_txt
		VAR_INPUT
			name 	: ^void;			//! <Variable Comment="Pointer to X509_NAME structure." Name="X509_NAME_add_entry_by_txt.name"/>
			field 	: ^void;			//! <Variable Comment="The field string represents the field name using OBJ_txt2obj(&lt;field&gt;, 0)." Name="X509_NAME_add_entry_by_txt.field"/>
			typ 	: DINT;			//! <Variable Comment="Field type.&#13;&#10;The use of string types such as MBSTRING_ASC or MBSTRING_UTF8 is strongly recommended for the type parameter. &#13;&#10;This allows the internal code to correctly determine the type of the field and to apply length checks according to the relevant standards. &#13;&#10;This is done using ASN1_STRING_set_by_NID().&#13;&#10;&#13;&#10;If instead an ASN1 type is used no checks are performed and the supplied data in bytes is used directly." Name="X509_NAME_add_entry_by_txt.typ"/>
			bytes 	: ^void;			//! <Variable Comment="Pointer to the field value to be added." Name="X509_NAME_add_entry_by_txt.bytes"/>
			len 	: DINT;			//! <Variable Comment="Length of the field value to be added.&#13;&#10;If &lt;len&gt; is -1 then the field length is calculated internally using strlen(&lt;bytes&gt;)." Name="X509_NAME_add_entry_by_txt.len"/>
			loc 	: DINT;			//! <Variable Comment="&lt;loc&gt; actually determines the index where the new entry is inserted: if it is -1 it is appended." Name="X509_NAME_add_entry_by_txt.loc"/>
			set 	: DINT;			//! <Variable Comment="&lt;set&gt; determines how the new type is added. If it is zero a new RDN is created.&#13;&#10;&#13;&#10;If &lt;set&gt; is -1 or 1 it is added to the previous or next RDN structure respectively. &#13;&#10;This will then be a multivalued RDN: since multivalues RDNs are very seldom used &lt;set&gt; is almost always set to zero." Name="X509_NAME_add_entry_by_txt.set"/>
		END_VAR
		VAR_OUTPUT
			RetVal (EAX) 	: DINT;			//! <Variable Comment="Returns 1 for success of 0 if an error occurred." Name="X509_NAME_add_entry_by_txt.RetVal"/>
		END_VAR;
				//! <Function Comment="X509_REVOKED_set_revocationDate() sets the revocation date of &lt;rx&gt; to &lt;tm&gt;. &#13;&#10;The supplied &lt;tm&gt; pointer is not used internally so it should be freed up after use.&#13;&#10;&#13;&#10;See also www.openssl.org/docs/man1.1.0/crypto/X509_REVOKED_set_revocationDate.html" Name="X509_REVOKED_set_revocationDate"/>
	FUNCTION __CDECL VIRTUAL GLOBAL X509_REVOKED_set_revocationDate
		VAR_INPUT
			rx 	: ^void;			//! <Variable Comment="Pointer to a X509_REVOKED structure." Name="X509_REVOKED_set_revocationDate.rx"/>
			tm 	: ^void;			//! <Variable Comment="Pointer to a ASN1_TIME structure holding the revocation date of &lt;rx&gt;.&#13;&#10;The supplied &lt;tm&gt; pointer is not used internally so it should be freed up after use." Name="X509_REVOKED_set_revocationDate.tm"/>
		END_VAR
		VAR_OUTPUT
			RetVal (EAX) 	: DINT;			//! <Variable Comment="Returns 1 for success and 0 for failure." Name="X509_REVOKED_set_revocationDate.RetVal"/>
		END_VAR;
				//! <Function Comment="Sets the issuer name of the CRL &lt;x&gt; to &lt;name&gt;.&#13;&#10;&#13;&#10;See also www.openssl.org/docs/man1.1.0/crypto/X509_CRL_set_issuer_name.html" Name="X509_CRL_set_issuer_name"/>
	FUNCTION __CDECL VIRTUAL GLOBAL X509_CRL_set_issuer_name
		VAR_INPUT
			x 	: ^void;			//! <Variable Comment="Pointer to X509_CRL structure holding a certificate revocation list (CRL)." Name="X509_CRL_set_issuer_name.x"/>
			name 	: ^void;			//! <Variable Comment="Pointer to X509_NAME structure holding the name to be set." Name="X509_CRL_set_issuer_name.name"/>
		END_VAR
		VAR_OUTPUT
			RetVal (EAX) 	: DINT;			//! <Variable Comment="Returns 1 for success and 0 for failure." Name="X509_CRL_set_issuer_name.RetVal"/>
		END_VAR;
				//! <Function Comment="X509_REVOKED_set_serialNumber() sets the serial number of &lt;x&gt; to &lt;serial&gt;. &#13;&#10;The supplied &lt;serial&gt; pointer is not used internally so it should be freed up after use.&#13;&#10;&#13;&#10;www.openssl.org/docs/man1.1.0/crypto/X509_REVOKED_set_serialNumber.html" Name="X509_REVOKED_set_serialNumber"/>
	FUNCTION __CDECL VIRTUAL GLOBAL X509_REVOKED_set_serialNumber
		VAR_INPUT
			x 	: ^void;			//! <Variable Comment="Pointer to a X509_REVOKED structure." Name="X509_REVOKED_set_serialNumber.x"/>
			serial 	: ^void;			//! <Variable Comment="Pointer to a ASN1_INTEGER structure holding the serial number to be set." Name="X509_REVOKED_set_serialNumber.serial"/>
		END_VAR
		VAR_OUTPUT
			RetVal (EAX) 	: DINT;			//! <Variable Comment="Returns 1 for success and 0 for failure." Name="X509_REVOKED_set_serialNumber.RetVal"/>
		END_VAR;
				//! <Function Comment="Releases the object and all pointers and sub-objects within it.&#13;&#10;&#13;&#10;See also www.openssl.org/docs/man1.1.0/crypto/X509_NAME_ENTRY_free.html" Name="X509_NAME_ENTRY_free"/>
	FUNCTION __CDECL VIRTUAL GLOBAL X509_NAME_ENTRY_free
		VAR_INPUT
			nex 	: ^void;			//! <Variable Comment="Pointer to a X509_NAME_ENTRY structure." Name="X509_NAME_ENTRY_free.nex"/>
		END_VAR;
				//! <Function Comment="Allocates an empty Certificate Revocation List (CRL). The CRL returned must be released by calling X509_CRL_free().&#13;&#10;&#13;&#10;See also www.openssl.org/docs/man1.1.0/crypto/X509_CRL_new.html" Name="X509_CRL_new"/>
	FUNCTION __CDECL VIRTUAL GLOBAL X509_CRL_new
		VAR_OUTPUT
			RetAddr (EAX) 	: ^void;			//! <Variable Comment="Returns a X509_CRL pointer to the newly created CRL or NULL on failure." Name="X509_CRL_new.RetAddr"/>
		END_VAR;
				//! <Function Comment="Releases the object and all pointers and sub-objects within it.&#13;&#10;&#13;&#10;See also www.openssl.org/docs/man1.1.0/crypto/X509_CRL_new.html" Name="X509_CRL_free"/>
	FUNCTION __CDECL VIRTUAL GLOBAL X509_CRL_free
		VAR_INPUT
			crl 	: ^void;			//! <Variable Comment="Pointer to X509_CRL structure holding a certificate revocation list (CRL)." Name="X509_CRL_free.crl"/>
		END_VAR;
				//! <Function Comment="Releases the object and all pointers and sub-objects within it.&#13;&#10;&#13;&#10;See also www.openssl.org/docs/man1.1.0/crypto/X509_CRL_new.html" Name="ASN1_TIME_free"/>
	FUNCTION __CDECL VIRTUAL GLOBAL ASN1_TIME_free
		VAR_INPUT
			mut 	: ^void;			//! <Variable Comment="Pointer to a ASN1_TIME structure." Name="ASN1_TIME_free.mut"/>
		END_VAR;
				//! <Function Comment="The ASN1_STRING object can represent a variety of ASN.1 built-in types. It can store a type and a value.&#13;&#10;&#13;&#10;The ASN1_INTEGER_new() function allocates and initializes an empty ASN1_STRING object.&#13;&#10;The object returned must be released by calling ASN1_INTEGER_free().&#13;&#10;&#13;&#10;See also https://users-cs.au.dk/sortie/sortix/release/nightly/man/man3/ASN1_INTEGER_new.3.html" Name="ASN1_INTEGER_new"/>
	FUNCTION __CDECL VIRTUAL GLOBAL ASN1_INTEGER_new
		VAR_OUTPUT
			RetAddr (EAX) 	: ^void;			//! <Variable Comment="Returns a ASN1_INTEGER pointer to the newly created object or NULL on failure." Name="ASN1_INTEGER_new.RetAddr"/>
		END_VAR;
				//! <Function Comment="Releases the object and all pointers and sub-objects within it.&#13;&#10;&#13;&#10;See also https://users-cs.au.dk/sortie/sortix/release/nightly/man/man3/ASN1_INTEGER_new.3.html" Name="ASN1_INTEGER_free"/>
	FUNCTION __CDECL VIRTUAL GLOBAL ASN1_INTEGER_free
		VAR_INPUT
			a 	: ^void;			//! <Variable Comment="Pointer to a ASN1_INTEGER object." Name="ASN1_INTEGER_free.a"/>
		END_VAR;
				//! <Function Comment="Allocates an empty object of the type X509_REVOKED. The object returned must be released by calling X509_REVOKED_free().&#13;&#10;&#13;&#10;See also www.openssl.org/docs/man1.1.0/crypto/X509_REVOKED_new.html" Name="X509_REVOKED_new"/>
	FUNCTION __CDECL VIRTUAL GLOBAL X509_REVOKED_new
		VAR_OUTPUT
			RetAddr (EAX) 	: ^void;			//! <Variable Comment="Returns a X509_REVOKED pointer to the newly created object or NULL on failure." Name="X509_REVOKED_new.RetAddr"/>
		END_VAR;
				//! <Function Comment="Releases the object and all pointers and sub-objects within it.&#13;&#10;&#13;&#10;See also www.openssl.org/docs/man1.1.0/crypto/X509_REVOKED_new.html" Name="X509_REVOKED_free"/>
	FUNCTION __CDECL VIRTUAL GLOBAL X509_REVOKED_free
		VAR_INPUT
			rx 	: ^void;			//! <Variable Comment="Pointer to a X509_REVOKED object." Name="X509_REVOKED_free.rx"/>
		END_VAR;
				//! <Function Comment="Writes the CRL &lt;x&gt; into the BIO &lt;bpx&gt; in PEM format.&#13;&#10;&#13;&#10;The PEM functions read or write structures in PEM format. In this sense PEM format is simply base64 encoded data surrounded by header lines.&#13;&#10;The X509_CRL functions process an X509 CRL using an X509_CRL structure.&#13;&#10;&#13;&#10;See also www.openssl.org/docs/man1.0.2/crypto/PEM_write_bio_X509_CRL.html" Name="PEM_write_bio_X509_CRL"/>
	FUNCTION __CDECL VIRTUAL GLOBAL PEM_write_bio_X509_CRL
		VAR_INPUT
			bpx 	: ^void;			//! <Variable Comment="Pointer to a BIO structure specifying the BIO to write to." Name="PEM_write_bio_X509_CRL.bpx"/>
			x 	: ^void;			//! <Variable Comment="Pointer to X509_CRL structure holding a certificate revocation list (CRL)." Name="PEM_write_bio_X509_CRL.x"/>
		END_VAR
		VAR_OUTPUT
			RetVal (EAX) 	: DINT;			//! <Variable Comment="Returns 1 for success or 0 for failure." Name="PEM_write_bio_X509_CRL.RetVal"/>
		END_VAR;
				//! <Function Comment="X509_cmp_time() compares the ASN1_TIME in &lt;sx&gt; with the time in &lt;tx&gt;. &#13;&#10;&#13;&#10;See also www.openssl.org/docs/man1.1.1/man3/X509_cmp_time.html" Name="X509_cmp_time"/>
	FUNCTION __CDECL VIRTUAL GLOBAL X509_cmp_time
		VAR_INPUT
			sx 	: ^void;			//! <Variable Comment="Pointer to a ASN1_TIME structure.&#13;&#10;&lt;sx&gt; must satisfy the ASN1_TIME format mandated by RFC 5280, i.e., its format must be either YYMMDDHHMMSSZ or YYYYMMDDHHMMSSZ (it&apos;s a literal Z at the end, meaning &quot;Zulu&quot;).&#13;&#10;" Name="X509_cmp_time.sx"/>
			tx 	: ^void;			//! <Variable Comment="Pointer to a time_t structure holding the number of seconds since the start of the Unix epoch: midnight UTC of January 1, 1970 (not counting leap seconds)." Name="X509_cmp_time.tx"/>
		END_VAR
		VAR_OUTPUT
			RetVal (EAX) 	: DINT;			//! <Variable Comment="Returns -1 if &lt;sx&gt; is earlier than, or equal to, &lt;tx&gt; and 1 otherwise. &#13;&#10;The method returns 0 on error." Name="X509_cmp_time.RetVal"/>
		END_VAR;
				//! <Function Comment="Returns the notBefore field of certificate &lt;x&gt;. The value returned is an internal pointer which must not be freed up after the call.&#13;&#10;&#13;&#10;See also www.openssl.org/docs/man1.1.0/crypto/X509_CRL_set1_lastUpdate.html" Name="X509_get_notBefore"/>
	FUNCTION __CDECL VIRTUAL GLOBAL X509_get_notBefore
		VAR_INPUT
			x 	: ^void;			//! <Variable Comment="Pointer to a X509 structure holding a certificate." Name="X509_get_notBefore.x"/>
		END_VAR
		VAR_OUTPUT
			RetAddr (EAX) 	: ^void;			//! <Variable Comment="Returns a pointer to an ASN1_TIME structure.&#13;&#10;Either YYMMDDHHMMSSZ or YYYYMMDDHHMMSSZ (it&apos;s a literal Z at the end, meaning &quot;Zulu&quot;)." Name="X509_get_notBefore.RetAddr"/>
		END_VAR;
				//! <Function Comment="Returns the notAfter field of certificate &lt;x&gt;. The value returned is an internal pointer which must not be freed up after the call.&#13;&#10;&#13;&#10;See also www.openssl.org/docs/man1.1.0/crypto/X509_CRL_set1_lastUpdate.html" Name="X509_get_notAfter"/>
	FUNCTION __CDECL VIRTUAL GLOBAL X509_get_notAfter
		VAR_INPUT
			x 	: ^void;			//! <Variable Comment="Pointer to a X509 structure holding a certificate." Name="X509_get_notAfter.x"/>
		END_VAR
		VAR_OUTPUT
			RetAddr (EAX) 	: ^void;			//! <Variable Comment="Returns a pointer to an ASN1_TIME structure.&#13;&#10;Either YYMMDDHHMMSSZ or YYYYMMDDHHMMSSZ (it&apos;s a literal Z at the end, meaning &quot;Zulu&quot;)." Name="X509_get_notAfter.RetAddr"/>
		END_VAR;
				//! <Function Comment="EVP_sha256(): the SHA-256 algorithm which produces a 160-bit output from a given input.&#13;&#10;SHA-256 (Secure Hash Algorithm 256) is a cryptographic hash function standardized in NIST FIPS 180-4.&#13;&#10;&#13;&#10;EVP_sha256() returns an EVP_MD structure for the SHA256 digest algorithm.&#13;&#10;&#13;&#10;See also www.openssl.org/docs/man1.0.2/crypto/EVP_sha256.html&#13;&#10;and       www.openssl.org/docs/man1.1.1/man3/EVP_sha256.html" Name="EVP_sha256"/>
	FUNCTION __CDECL VIRTUAL GLOBAL EVP_sha256
		VAR_OUTPUT
			RetAddr (EAX) 	: ^void;			//! <Variable Comment="Pointer to an EVP_MD structure that contains the implementation of the symmetric cipher." Name="EVP_sha256.RetAddr"/>
		END_VAR;
				//! <Function Comment="SHA-256 (Secure Hash Algorithm) is a cryptographic hash function with a 160 bit output.&#13;&#10;&#13;&#10;SHA256() computes the SHA-256 message digest of the &lt;n_val&gt; bytes at &lt;d_addr&gt; and places it in &lt;md&gt; (which must have space for SHA256_DIGEST_LENGTH).&#13;&#10;If &lt;md&gt; is NULL, the digest is placed in a static array. Note: setting &lt;md&gt; to NULL is not thread safe.&#13;&#10;&#13;&#10;See also www.openssl.org/docs/man1.0.2/crypto/SHA256.html" Name="SHA256"/>
	FUNCTION __CDECL VIRTUAL GLOBAL SHA256
		VAR_INPUT
			d_addr 	: ^USINT;			//! <Variable Comment="Pointer to input buffer." Name="SHA256.d_addr"/>
			n_val 	: DINT;			//! <Variable Comment="Length of the input buffer in bytes." Name="SHA256.n_val"/>
			md 	: ^USINT;			//! <Variable Comment="Pointer to the SHA-256 message digest buffer (&lt;md&gt; must have space for SHA256_DIGEST_LENGTH). &#13;&#10;If &lt;md&gt; is NULL, the digest is placed in a static array (WARNING: not thread-safe)." Name="SHA256.md"/>
		END_VAR
		VAR_OUTPUT
			RetAddr (EAX) 	: ^USINT;			//! <Variable Comment="Returns a pointer to the hash value." Name="SHA256.RetAddr"/>
		END_VAR;
				//! <Function Comment="Writes data from buffer to BIO b." Name="BIO_write"/>
	FUNCTION __CDECL VIRTUAL GLOBAL BIO_write
		VAR_INPUT
			b 	: ^void;			//! <Variable Comment="Pointer to BIO structure." Name="BIO_write.b"/>
			data 	: ^void;			//! <Variable Comment="Pointer to the data buffer." Name="BIO_write.data"/>
			len 	: DINT;			//! <Variable Comment="Number of bytes to write from data to BIO b." Name="BIO_write.len"/>
		END_VAR
		VAR_OUTPUT
			RetVal (EAX) 	: DINT;			//! <Variable Comment="Returns -2 if the &quot;write&quot; operation is not implemented by the BIO or -1 on other errors. Otherwise it returns the number of bytes written. This may be 0 if the BIO b is NULL or dlen &lt;= 0." Name="BIO_write.RetVal"/>
		END_VAR;
				//! <Function Comment="Reads an RSA public key using an RSA structure." Name="PEM_read_bio_RSA_PUBKEY"/>
	FUNCTION __CDECL VIRTUAL GLOBAL PEM_read_bio_RSA_PUBKEY
		VAR_INPUT
			b 	: ^void;			//! <Variable Comment="Specifies the BIO to read from." Name="PEM_read_bio_RSA_PUBKEY.b"/>
			x 	: ^pVoid;			//! <Variable Comment="If x is NULL then the parameter is ignored. &#13;&#10;If x is not NULL but *x is NULL then the structure returned will be written to *x. &#13;&#10;If neither x nor *x is NULL then an attempt is made to reuse the structure at *x. &#13;&#10;Irrespective of the value of x a pointer to the structure is always returned (or NULL if an error occurred)." Name="PEM_read_bio_RSA_PUBKEY.x"/>
			cb 	: ^void;			//! <Variable Comment="The cb argument is the callback to use when querying for the pass phrase used for encrypted PEM structures." Name="PEM_read_bio_RSA_PUBKEY.cb"/>
			u 	: ^void;			//! <Variable Comment="If the cb parameters is set to NULL and the u parameter is not NULL then the u parameter is interpreted as a null terminated string to use as the passphrase. &#13;&#10;If both cb and u are NULL then the default callback routine is used." Name="PEM_read_bio_RSA_PUBKEY.u"/>
		END_VAR
		VAR_OUTPUT
			RetAddr (EAX) 	: ^void;			//! <Variable Comment="Returns a pointer to an RSA structure." Name="PEM_read_bio_RSA_PUBKEY.RetAddr"/>
		END_VAR;
				//! <Function Comment="Initializes a SHA512_CTX structure." Name="SHA512_Init"/>
	FUNCTION __CDECL VIRTUAL GLOBAL SHA512_Init
		VAR_INPUT
			c 	: ^void;			//! <Variable Comment="Pointer to the SHA512_CTX structure." Name="SHA512_Init.c"/>
		END_VAR
		VAR_OUTPUT
			RetVal (EAX) 	: DINT;			//! <Variable Comment="Return 1 for success, 0 otherwise." Name="SHA512_Init.RetVal"/>
		END_VAR;
				//! <Function Comment="Can be called repeatedly with chunks of the message to be hashed (len bytes at data)." Name="SHA512_Update"/>
	FUNCTION __CDECL VIRTUAL GLOBAL SHA512_Update
		VAR_INPUT
			c 	: ^void;			//! <Variable Comment="Pointer to the SHA512_CTX structure." Name="SHA512_Update.c"/>
			data 	: ^void;			//! <Variable Comment="Pointer to the data buffer." Name="SHA512_Update.data"/>
			len 	: DINT;			//! <Variable Comment="Data buffer length." Name="SHA512_Update.len"/>
		END_VAR
		VAR_OUTPUT
			RetVal (EAX) 	: DINT;			//! <Variable Comment="Return 1 for success, 0 otherwise." Name="SHA512_Update.RetVal"/>
		END_VAR;
				//! <Function Comment="Places the message digest in md, which must have space for SHA512_DIGEST_LENGTH == 64 bytes of output, and erases the SHA512_CTX." Name="SHA512_Final"/>
	FUNCTION __CDECL VIRTUAL GLOBAL SHA512_Final
		VAR_INPUT
			md 	: ^USINT;			//! <Variable Comment="Pointer to the SHA-512 message digest buffer (&lt;md&gt; must have space for SHA512_DIGEST_LENGTH). &#13;&#10;If &lt;md&gt; is NULL, the digest is placed in a static array (WARNING: not thread-safe)." Name="SHA512_Final.md"/>
			c 	: ^void;			//! <Variable Comment="Pointer to the SHA512_CTX structure." Name="SHA512_Final.c"/>
		END_VAR
		VAR_OUTPUT
			RetVal (EAX) 	: DINT;			//! <Variable Comment="Return 1 for success, 0 otherwise." Name="SHA512_Final.RetVal"/>
		END_VAR;
				//! <Function Comment="SHA-512 (Secure Hash Algorithm) is a cryptographic hash function.&#13;&#10;&#13;&#10;SHA512() computes the SHA-512 message digest of the &lt;n_val&gt; bytes at &lt;d_addr&gt; and places it in &lt;md&gt; (which must have space for SHA512_DIGEST_LENGTH).&#13;&#10;If &lt;md&gt; is NULL, the digest is placed in a static array. Note: setting &lt;md&gt; to NULL is not thread safe." Name="SHA512"/>
	FUNCTION __CDECL VIRTUAL GLOBAL SHA512
		VAR_INPUT
			d_addr 	: ^USINT;			//! <Variable Comment="Pointer to input buffer." Name="SHA512.d_addr"/>
			n_val 	: DINT;			//! <Variable Comment="Length of the input buffer in bytes." Name="SHA512.n_val"/>
			md 	: ^USINT;			//! <Variable Comment="Pointer to the SHA-512 message digest buffer (&lt;md&gt; must have space for SHA512_DIGEST_LENGTH). &#13;&#10;If &lt;md&gt; is NULL, the digest is placed in a static array (WARNING: not thread-safe)." Name="SHA512.md"/>
		END_VAR
		VAR_OUTPUT
			RetAddr (EAX) 	: ^USINT;			//! <Variable Comment="Returns a pointer to the hash value." Name="SHA512.RetAddr"/>
		END_VAR;
  //Tables:
	FUNCTION @STD
		VAR_OUTPUT
			ret_code	: CONFSTATES;
		END_VAR;
	FUNCTION GLOBAL TAB @CT_;
END_CLASS;

#include <Rtos_interfaces.h> // we need this for the SysCIL functions
#include "..\..\Source\code\OsiBaseNew.h"

// This variable has to be global to allow for calls to OpenSSL CIL API
// functions from C code without the C programmer needing to call OS_CILGet
// explicitly. In such a case the CIL API functions are called via C macros
// defined in lsl_c_openssl.h.
VAR_GLOBAL
  lsl_openssl   : ^_OpenSSL::LSL_OPENSSL; //Used for compatibility of previous versions
  _lsl_openssl  : ^_OpenSSL::LSL_OPENSSL; //Used for function calls in c
END_VAR

VAR_PRIVATE
   API_Version:UDINT;
END_VAR

FUNCTION VIRTUAL GLOBAL _OpenSSL::GetVersion
	VAR_OUTPUT
		ret0 	: UDINT;
	END_VAR
   ret0 := API_Version;
END_FUNCTION

// Disable 'Parameter '...' is never used' warnings
#pragma warning (disable:73)
// Dummy functions

FUNCTION __CDECL _OpenSSL_DummyInt
VAR_OUTPUT
  dRC      : DINT;
END_VAR
  dRC := OpenSSL_ERR_NO_INTERFACE;
END_FUNCTION

FUNCTION __CDECL _OpenSSL_DummyPtr
VAR_OUTPUT
  pOutput  : pVoid;
END_VAR
  pOutput := nil;
END_FUNCTION

FUNCTION __CDECL _OpenSSL_DummyVoid

END_FUNCTION

#pragma warning (default:73)
// End of Dummy functions

FUNCTION _OpenSSL::_OpenSSL
	VAR_OUTPUT
		ret_code 	: ConfStates;
	END_VAR

VAR
	aMeths			: ARRAY[0..USER_CNT__OpenSSL] OF ^void;
	retv    		: SYS_ERROR;
END_VAR

	retv := OS_CILGet(INTERFACE_OPENSSL, #lsl_openssl);
	_lsl_openssl := lsl_openssl;

	if retv <> SYS_ERR_NONE then

	  TRACE("ERROR: OPENSSL interface not available with this version/platform");

    API_Version := 0;

    aMeths[0]  := #GetVersion();
    aMeths[1]  := #_OpenSSL_DummyPtr();
		aMeths[2]  := #_OpenSSL_DummyPtr();
		aMeths[3]  := #_OpenSSL_DummyInt();
		aMeths[4]  := #_OpenSSL_DummyPtr();
		aMeths[5]  := #_OpenSSL_DummyPtr();
		aMeths[6]  := #_OpenSSL_DummyInt();
		aMeths[7]  := #_OpenSSL_DummyVoid();
		aMeths[8]  := #_OpenSSL_DummyVoid();
 	  aMeths[9]  := #_OpenSSL_DummyPtr();
    aMeths[10] := #_OpenSSL_DummyVoid();
    aMeths[11] := #_OpenSSL_DummyVoid();
    aMeths[12] := #_OpenSSL_DummyInt();
		aMeths[13] := #_OpenSSL_DummyVoid();
		aMeths[14] := #_OpenSSL_DummyVoid();
		aMeths[15] := #_OpenSSL_DummyVoid();
		aMeths[16] := #_OpenSSL_DummyVoid();
    aMeths[17] := #_OpenSSL_DummyInt();
		aMeths[18] := #_OpenSSL_DummyInt();
		aMeths[19] := #_OpenSSL_DummyVoid();
    aMeths[20] := #_OpenSSL_DummyPtr();
	  aMeths[21] := #_OpenSSL_DummyPtr();
		aMeths[22] := #_OpenSSL_DummyVoid();
		aMeths[23] := #_OpenSSL_DummyInt();
		aMeths[24] := #_OpenSSL_DummyPtr();
		aMeths[25] := #_OpenSSL_DummyInt();
		aMeths[26] := #_OpenSSL_DummyPtr();
		aMeths[27] := #_OpenSSL_DummyInt();
		aMeths[28] := #_OpenSSL_DummyInt();
		aMeths[29] := #_OpenSSL_DummyPtr();
		aMeths[30] := #_OpenSSL_DummyPtr();
		aMeths[31] := #_OpenSSL_DummyPtr();
		aMeths[32] := #_OpenSSL_DummyVoid();
		aMeths[33] := #_OpenSSL_DummyPtr();
		aMeths[34] := #_OpenSSL_DummyPtr();
		aMeths[35] := #_OpenSSL_DummyPtr();
		aMeths[36] := #_OpenSSL_DummyInt();
		aMeths[37] := #_OpenSSL_DummyVoid();
		aMeths[38] := #_OpenSSL_DummyPtr();
		aMeths[39] := #_OpenSSL_DummyVoid();
		aMeths[40] := #_OpenSSL_DummyInt();
		aMeths[41] := #_OpenSSL_DummyInt();
		aMeths[42] := #_OpenSSL_DummyInt();
		aMeths[43] := #_OpenSSL_DummyInt();
		aMeths[44] := #_OpenSSL_DummyInt();
		aMeths[45] := #_OpenSSL_DummyInt();
		aMeths[46] := #_OpenSSL_DummyInt();
		aMeths[47] := #_OpenSSL_DummyPtr();
		aMeths[48] := #_OpenSSL_DummyInt();
		aMeths[49] := #_OpenSSL_DummyInt();
		aMeths[50] := #_OpenSSL_DummyPtr();
		aMeths[51] := #_OpenSSL_DummyInt();
		aMeths[52] := #_OpenSSL_DummyPtr();
		aMeths[53] := #_OpenSSL_DummyInt();
		aMeths[54] := #_OpenSSL_DummyVoid();
		aMeths[55] := #_OpenSSL_DummyPtr();
		aMeths[56] := #_OpenSSL_DummyInt();
		aMeths[57] := #_OpenSSL_DummyPtr();
		aMeths[58] := #_OpenSSL_DummyPtr();
		aMeths[59] := #_OpenSSL_DummyInt();
		aMeths[60] := #_OpenSSL_DummyInt();
		aMeths[61] := #_OpenSSL_DummyPtr();
		aMeths[62] := #_OpenSSL_DummyInt();
		aMeths[63] := #_OpenSSL_DummyInt();
		aMeths[64] := #_OpenSSL_DummyPtr();
		aMeths[65] := #_OpenSSL_DummyVoid();
		aMeths[66] := #_OpenSSL_DummyInt();
		aMeths[67] := #_OpenSSL_DummyVoid();
		aMeths[68] := #_OpenSSL_DummyInt();
		aMeths[69] := #_OpenSSL_DummyPtr();
		aMeths[70] := #_OpenSSL_DummyPtr();
		aMeths[71] := #_OpenSSL_DummyPtr();
		aMeths[72] := #_OpenSSL_DummyInt();
    aMeths[73] := #_OpenSSL_DummyPtr();
    aMeths[74] := #_OpenSSL_DummyInt();
    aMeths[75] := #_OpenSSL_DummyInt();
    aMeths[76] := #_OpenSSL_DummyPtr();
    aMeths[77] := #_OpenSSL_DummyInt();
    aMeths[78] := #_OpenSSL_DummyPtr();
    aMeths[79] := #_OpenSSL_DummyInt();
    aMeths[80] := #_OpenSSL_DummyInt();
    aMeths[81] := #_OpenSSL_DummyPtr();
    aMeths[82] := #_OpenSSL_DummyInt();
    aMeths[83] := #_OpenSSL_DummyPtr();
    aMeths[84] := #_OpenSSL_DummyVoid();
    aMeths[85] := #_OpenSSL_DummyInt();
    aMeths[86] := #_OpenSSL_DummyPtr();
    aMeths[87] := #_OpenSSL_DummyInt();
    aMeths[88] := #_OpenSSL_DummyInt();
    aMeths[89] := #_OpenSSL_DummyPtr();
    aMeths[90] := #_OpenSSL_DummyInt();
    aMeths[91] := #_OpenSSL_DummyPtr();
    aMeths[92] := #_OpenSSL_DummyInt();
    aMeths[93] := #_OpenSSL_DummyInt();
    aMeths[94] := #_OpenSSL_DummyPtr();
    aMeths[95] := #_OpenSSL_DummyInt();
    aMeths[96] := #_OpenSSL_DummyPtr();
    aMeths[97] := #_OpenSSL_DummyInt();
    aMeths[98] := #_OpenSSL_DummyInt();
    aMeths[99] := #_OpenSSL_DummyPtr();
    aMeths[100] := #_OpenSSL_DummyInt();
    aMeths[101] := #_OpenSSL_DummyPtr();
    aMeths[102] := #_OpenSSL_DummyPtr();
    aMeths[103] := #_OpenSSL_DummyInt();
    aMeths[104] := #_OpenSSL_DummyInt();
    aMeths[105] := #_OpenSSL_DummyPtr();
    aMeths[106] := #_OpenSSL_DummyPtr();
    aMeths[107] := #_OpenSSL_DummyInt();
    aMeths[108] := #_OpenSSL_DummyPtr();
    aMeths[109] := #_OpenSSL_DummyInt();
    aMeths[110] := #_OpenSSL_DummyInt();
    aMeths[111] := #_OpenSSL_DummyInt();
    aMeths[112] := #_OpenSSL_DummyInt();
    aMeths[113] := #_OpenSSL_DummyInt();
    aMeths[114] := #_OpenSSL_DummyInt();
    aMeths[115] := #_OpenSSL_DummyInt();
    aMeths[116] := #_OpenSSL_DummyInt();
    aMeths[117] := #_OpenSSL_DummyInt();
    aMeths[118] := #_OpenSSL_DummyInt();
    aMeths[119] := #_OpenSSL_DummyInt();
    aMeths[120] := #_OpenSSL_DummyInt();
    aMeths[121] := #_OpenSSL_DummyVoid();
    aMeths[122] := #_OpenSSL_DummyPtr();
    aMeths[123] := #_OpenSSL_DummyVoid();
    aMeths[124] := #_OpenSSL_DummyVoid();
    aMeths[125] := #_OpenSSL_DummyPtr();
    aMeths[126] := #_OpenSSL_DummyVoid();
    aMeths[127] := #_OpenSSL_DummyPtr();
    aMeths[128] := #_OpenSSL_DummyVoid();
    aMeths[129] := #_OpenSSL_DummyInt();
    aMeths[130] := #_OpenSSL_DummyInt();
    aMeths[131] := #_OpenSSL_DummyPtr();
    aMeths[132] := #_OpenSSL_DummyPtr();
    aMeths[133] := #_OpenSSL_DummyPtr();
    aMeths[134] := #_OpenSSL_DummyPtr();

  else
    API_Version := lsl_openssl^.udVersion;

    aMeths[0]  := #GetVersion();
    aMeths[1]  := lsl_openssl^.d2i_X509;
		aMeths[2]  := lsl_openssl^.X509_get_subject_name;
		aMeths[3]  := lsl_openssl^.X509_NAME_get_index_by_NID;
		aMeths[4]  := lsl_openssl^.X509_NAME_get_entry;
		aMeths[5]  := lsl_openssl^.X509_NAME_ENTRY_get_data;
		aMeths[6]  := lsl_openssl^.ASN1_STRING_to_UTF8;
		aMeths[7]  := lsl_openssl^.OPENSSL_free;
		aMeths[8]  := lsl_openssl^.X509_free;
		aMeths[9]  := lsl_openssl^.SSLeay_version;
		aMeths[10] := lsl_openssl^.OpenSSL_add_all_algorithms;
		aMeths[11] := lsl_openssl^.ERR_load_crypto_strings;
		aMeths[12] := lsl_openssl^.X509_STORE_CTX_get_ex_new_index;
		aMeths[13] := lsl_openssl^.EVP_cleanup;
		aMeths[14] := lsl_openssl^.CRYPTO_cleanup_all_ex_data;
		aMeths[15] := lsl_openssl^.ERR_remove_state;
		aMeths[16] := lsl_openssl^.ERR_free_strings;
		aMeths[17] := lsl_openssl^.AES_set_encrypt_key;
		aMeths[18] := lsl_openssl^.AES_set_decrypt_key;
		aMeths[19] := lsl_openssl^.AES_cbc_encrypt;

		aMeths[20] := lsl_openssl^.EVP_sha1;
		aMeths[21] := lsl_openssl^.HMAC;
		aMeths[22] := lsl_openssl^.X509_STORE_free;
		aMeths[23] := lsl_openssl^.X509_STORE_add_cert;
		aMeths[24] := lsl_openssl^.SHA1;

		aMeths[25] := lsl_openssl^.RAND_bytes;

		aMeths[26] := lsl_openssl^.RSA_generate_key;
		aMeths[27] := lsl_openssl^.i2d_RSAPublicKey;
		aMeths[28] := lsl_openssl^.i2d_RSAPrivateKey;
		aMeths[29] := lsl_openssl^.d2i_RSAPrivateKey;
		aMeths[30] := lsl_openssl^.d2i_PublicKey;
		aMeths[31] := lsl_openssl^.d2i_PrivateKey;
		aMeths[32] := lsl_openssl^.RSA_free;
		aMeths[33] := lsl_openssl^.BIO_new_file;
		aMeths[34] := lsl_openssl^.PEM_read_bio_PrivateKey;
		aMeths[35] := lsl_openssl^.d2i_PKCS12_bio;
		aMeths[36] := lsl_openssl^.PKCS12_parse;
		aMeths[37] := lsl_openssl^.PKCS12_free;
		aMeths[38] := lsl_openssl^.EVP_PKEY_get1_RSA;
		aMeths[39] := lsl_openssl^.EVP_PKEY_free;
		aMeths[40] := lsl_openssl^.BIO_free;
		aMeths[41] := lsl_openssl^.PEM_write_bio_RSAPrivateKey;
		aMeths[42] := lsl_openssl^.RSA_size;
		aMeths[43] := lsl_openssl^.RSA_public_encrypt;
		aMeths[44] := lsl_openssl^.RSA_private_decrypt;
		aMeths[45] := lsl_openssl^.RSA_sign;
		aMeths[46] := lsl_openssl^.ERR_get_error;
		aMeths[47] := lsl_openssl^.ERR_error_string;
		aMeths[48] := lsl_openssl^.RSA_verify;

		aMeths[49] := lsl_openssl^.OBJ_txt2nid;
		aMeths[50] := lsl_openssl^.X509_NAME_ENTRY_create_by_NID;
		aMeths[51] := lsl_openssl^.X509_NAME_add_entry;
		aMeths[52] := lsl_openssl^.X509V3_EXT_conf;
		aMeths[53] := lsl_openssl^.X509_add_ext;
		aMeths[54] := lsl_openssl^.X509_EXTENSION_free;
		aMeths[55] := lsl_openssl^.X509_new;
		aMeths[56] := lsl_openssl^.X509_set_version;
		aMeths[57] := lsl_openssl^.X509_get_serialNumber;
		aMeths[58] := lsl_openssl^.OPENSSL_Realloc;
		aMeths[59] := lsl_openssl^.ASN1_INTEGER_set;
		aMeths[60] := lsl_openssl^.X509_set_pubkey;
		aMeths[61] := lsl_openssl^.X509_NAME_new;
		aMeths[62] := lsl_openssl^.X509_set_subject_name;
		aMeths[63] := lsl_openssl^.X509_set_issuer_name;
		aMeths[64] := lsl_openssl^.X509_gmtime_adj;
		aMeths[65] := lsl_openssl^.X509V3_set_ctx;
		aMeths[66] := lsl_openssl^.X509_sign;
		aMeths[67] := lsl_openssl^.X509_NAME_free;
		aMeths[68] := lsl_openssl^.i2d_X509_bio;
		aMeths[69] := lsl_openssl^.d2i_X509_bio;
		aMeths[70] := lsl_openssl^.PEM_read_bio_X509;
		aMeths[71] := lsl_openssl^.X509_get_pubkey;
		aMeths[72] := lsl_openssl^.OBJ_obj2nid;

    if API_Version >= 2 then

      aMeths[73] := lsl_openssl^.BIO_new;
      aMeths[74] := lsl_openssl^.i2d_X509;
      aMeths[75] := lsl_openssl^.X509_verify;
      aMeths[76] := lsl_openssl^.X509_STORE_new;
      aMeths[77] := lsl_openssl^.CRYPTO_add_lock;
      aMeths[78] := lsl_openssl^.X509_LOOKUP_file;
      aMeths[79] := lsl_openssl^.X509_LOOKUP_ctrl;
      aMeths[80] := lsl_openssl^.X509_verify_cert;
      aMeths[81] := lsl_openssl^.X509_NAME_oneline;
      aMeths[82] := lsl_openssl^.X509_load_crl_file;
      aMeths[83] := lsl_openssl^.X509_STORE_CTX_new;
      aMeths[84] := lsl_openssl^.X509_STORE_CTX_free;
      aMeths[85] := lsl_openssl^.X509_STORE_CTX_init;
      aMeths[86] := lsl_openssl^.X509_get_issuer_name;
      aMeths[87] := lsl_openssl^.X509_LOOKUP_hash_dir;
      aMeths[88] := lsl_openssl^.X509_STORE_set_flags;
      aMeths[89] := lsl_openssl^.X509_STORE_add_lookup;
      aMeths[90]:= lsl_openssl^.X509_STORE_set_default_paths;
      aMeths[91] := lsl_openssl^.X509_STORE_CTX_get_ex_data;
      aMeths[92]:= lsl_openssl^.X509_STORE_CTX_set_ex_data;
      aMeths[93] := lsl_openssl^.X509_STORE_CTX_get_error;
      aMeths[94] := lsl_openssl^.X509_STORE_CTX_get_current_cert;
      aMeths[95] := lsl_openssl^.X509_STORE_CTX_get_error_depth;
      aMeths[96] := lsl_openssl^.X509_verify_cert_error_string;
      aMeths[97] := lsl_openssl^.i2d_PublicKey;
      aMeths[98] := lsl_openssl^.EVP_PKEY_type;
      aMeths[99] := lsl_openssl^.CRYPTO_realloc;
      aMeths[100] := lsl_openssl^.BIO_ctrl;
      aMeths[101] := lsl_openssl^.BIO_s_mem;
      aMeths[102] := lsl_openssl^.BIO_s_file;
      aMeths[103] := lsl_openssl^.X509_get_ext;
      aMeths[104] := lsl_openssl^.EVP_PKEY_cmp;
      aMeths[105] := lsl_openssl^.EVP_PKEY_new;
      aMeths[106] := lsl_openssl^.ASN1_TIME_set;
      aMeths[107] := lsl_openssl^.X509_CRL_sign;
      aMeths[108] := lsl_openssl^.X509_PUBKEY_get;
      aMeths[109] := lsl_openssl^.EVP_PKEY_assign;
      aMeths[110] := lsl_openssl^.X509V3_EXT_print;
      aMeths[111] := lsl_openssl^.X509_get_ext_by_NID;
      aMeths[112] := lsl_openssl^.X509_CRL_set_version;
      aMeths[113] := lsl_openssl^.X509_CRL_add0_revoked;
      aMeths[114] := lsl_openssl^.X509_CRL_add1_ext_i2d;
      aMeths[115] := lsl_openssl^.X509_CRL_set_lastUpdate;
      aMeths[116] := lsl_openssl^.X509_CRL_set_nextUpdate;
      aMeths[117] := lsl_openssl^.X509_NAME_add_entry_by_txt;
      aMeths[118] := lsl_openssl^.X509_REVOKED_set_revocationDate;
      aMeths[119] := lsl_openssl^.X509_CRL_set_issuer_name;
      aMeths[120] := lsl_openssl^.X509_REVOKED_set_serialNumber;
      aMeths[121] := lsl_openssl^.X509_NAME_ENTRY_free;
      aMeths[122] := lsl_openssl^.X509_CRL_new;
      aMeths[123] := lsl_openssl^.X509_CRL_free;
      aMeths[124] := lsl_openssl^.ASN1_TIME_free;
      aMeths[125] := lsl_openssl^.ASN1_INTEGER_new;
      aMeths[126] := lsl_openssl^.ASN1_INTEGER_free;
      aMeths[127] := lsl_openssl^.X509_REVOKED_new;
      aMeths[128] := lsl_openssl^.X509_REVOKED_free;
      aMeths[129] := lsl_openssl^.PEM_write_bio_X509_CRL;
      aMeths[130] := lsl_openssl^.X509_cmp_time;

    else

      aMeths[73] := #_OpenSSL_DummyPtr();
      aMeths[74] := #_OpenSSL_DummyInt();
      aMeths[75] := #_OpenSSL_DummyInt();
      aMeths[76] := #_OpenSSL_DummyPtr();
      aMeths[77] := #_OpenSSL_DummyInt();
      aMeths[78] := #_OpenSSL_DummyPtr();
      aMeths[79] := #_OpenSSL_DummyInt();
      aMeths[80] := #_OpenSSL_DummyInt();
      aMeths[81] := #_OpenSSL_DummyPtr();
      aMeths[82] := #_OpenSSL_DummyInt();
      aMeths[83] := #_OpenSSL_DummyPtr();
      aMeths[84] := #_OpenSSL_DummyVoid();
      aMeths[85] := #_OpenSSL_DummyInt();
      aMeths[86] := #_OpenSSL_DummyPtr();
      aMeths[87] := #_OpenSSL_DummyInt();
      aMeths[88] := #_OpenSSL_DummyInt();
      aMeths[89] := #_OpenSSL_DummyPtr();
      aMeths[90] := #_OpenSSL_DummyInt();
      aMeths[91] := #_OpenSSL_DummyPtr();
      aMeths[92] := #_OpenSSL_DummyInt();
      aMeths[93] := #_OpenSSL_DummyInt();
      aMeths[94] := #_OpenSSL_DummyPtr();
      aMeths[95] := #_OpenSSL_DummyInt();
      aMeths[96] := #_OpenSSL_DummyPtr();
      aMeths[97] := #_OpenSSL_DummyInt();
      aMeths[98] := #_OpenSSL_DummyInt();
      aMeths[99] := #_OpenSSL_DummyPtr();
      aMeths[100] := #_OpenSSL_DummyInt();
      aMeths[101] := #_OpenSSL_DummyPtr();
      aMeths[102] := #_OpenSSL_DummyPtr();
      aMeths[103] := #_OpenSSL_DummyInt();
      aMeths[104] := #_OpenSSL_DummyInt();
      aMeths[105] := #_OpenSSL_DummyPtr();
      aMeths[106] := #_OpenSSL_DummyPtr();
      aMeths[107] := #_OpenSSL_DummyInt();
      aMeths[108] := #_OpenSSL_DummyPtr();
      aMeths[109] := #_OpenSSL_DummyInt();
      aMeths[110] := #_OpenSSL_DummyInt();
      aMeths[111] := #_OpenSSL_DummyInt();
      aMeths[112] := #_OpenSSL_DummyInt();
      aMeths[113] := #_OpenSSL_DummyInt();
      aMeths[114] := #_OpenSSL_DummyInt();
      aMeths[115] := #_OpenSSL_DummyInt();
      aMeths[116] := #_OpenSSL_DummyInt();
      aMeths[117] := #_OpenSSL_DummyInt();
      aMeths[118] := #_OpenSSL_DummyInt();
      aMeths[119] := #_OpenSSL_DummyInt();
      aMeths[120] := #_OpenSSL_DummyInt();
      aMeths[121] := #_OpenSSL_DummyVoid();
      aMeths[122] := #_OpenSSL_DummyPtr();
      aMeths[123] := #_OpenSSL_DummyVoid();
      aMeths[124] := #_OpenSSL_DummyVoid();
      aMeths[125] := #_OpenSSL_DummyPtr();
      aMeths[126] := #_OpenSSL_DummyVoid();
      aMeths[127] := #_OpenSSL_DummyPtr();
      aMeths[128] := #_OpenSSL_DummyVoid();
      aMeths[129] := #_OpenSSL_DummyInt();
      aMeths[130] := #_OpenSSL_DummyInt();

    end_if;

    if API_Version >= 3 then

      aMeths[131] := lsl_openssl^.X509_get_notBefore;
      aMeths[132] := lsl_openssl^.X509_get_notAfter;

    else

      aMeths[131] := #_OpenSSL_DummyPtr();
      aMeths[132] := #_OpenSSL_DummyPtr();

    end_if;

    if API_Version >= 4 then

      aMeths[133] := lsl_openssl^.EVP_sha256;
      aMeths[134] := lsl_openssl^.SHA256;

    else

      aMeths[133] := #_OpenSSL_DummyPtr();
      aMeths[134] := #_OpenSSL_DummyPtr();

    end_if;

    if API_Version >= 5 then

      aMeths[135] := lsl_openssl^.BIO_write;
      aMeths[136] := lsl_openssl^.PEM_read_bio_RSA_PUBKEY;
      aMeths[137] := lsl_openssl^.SHA512_Init;
      aMeths[138] := lsl_openssl^.SHA512_Update;
      aMeths[139] := lsl_openssl^.SHA512_Final;
      aMeths[140] := lsl_openssl^.SHA512;

    else

      aMeths[135] := #_OpenSSL_DummyInt();
      aMeths[136] := #_OpenSSL_DummyPtr();
      aMeths[137] := #_OpenSSL_DummyInt();
      aMeths[138] := #_OpenSSL_DummyInt();
      aMeths[139] := #_OpenSSL_DummyInt();
      aMeths[140] := #_OpenSSL_DummyPtr();

    end_if;

	end_if;

  // Hier das Array mit weiteren Zeigern auf API-Funktionen initialisieren ...
  ret_code  := InitOsiM_new(#aMeths[0]$void, USER_CNT__OpenSSL);

END_FUNCTION
